FUNCTION_BLOCK TestingSequence1 (* Composite Function Block Type *)
  (* Standard: 61499-2 *)
  (* Version 0.0, 7/2/2026, template *)
  PACKAGE Main;
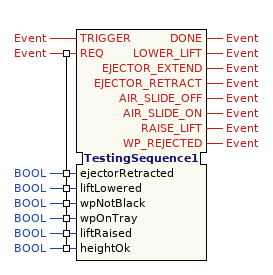
  EVENT_INPUT
    TRIGGER; (* Initialization Request *)
    REQ WITH ejectorRetracted, liftLowered, wpNotBlack, wpOnTray, liftRaised, heightOk; (* Normal Execution Request *)
  END_EVENT
  EVENT_OUTPUT
    DONE; (* Initialization Confirm *)
    LOWER_LIFT; (* Execution Confirmation *)
    EJECTOR_EXTEND;
    EJECTOR_RETRACT;
    AIR_SLIDE_OFF;
    AIR_SLIDE_ON;
    RAISE_LIFT;
    WP_REJECTED;
  END_EVENT
  VAR_INPUT
    ejectorRetracted : BOOL; (* Input event qualifier *)
    liftLowered : BOOL;
    wpNotBlack : BOOL;
    wpOnTray : BOOL;
    liftRaised : BOOL;
    heightOk : BOOL;
  END_VAR
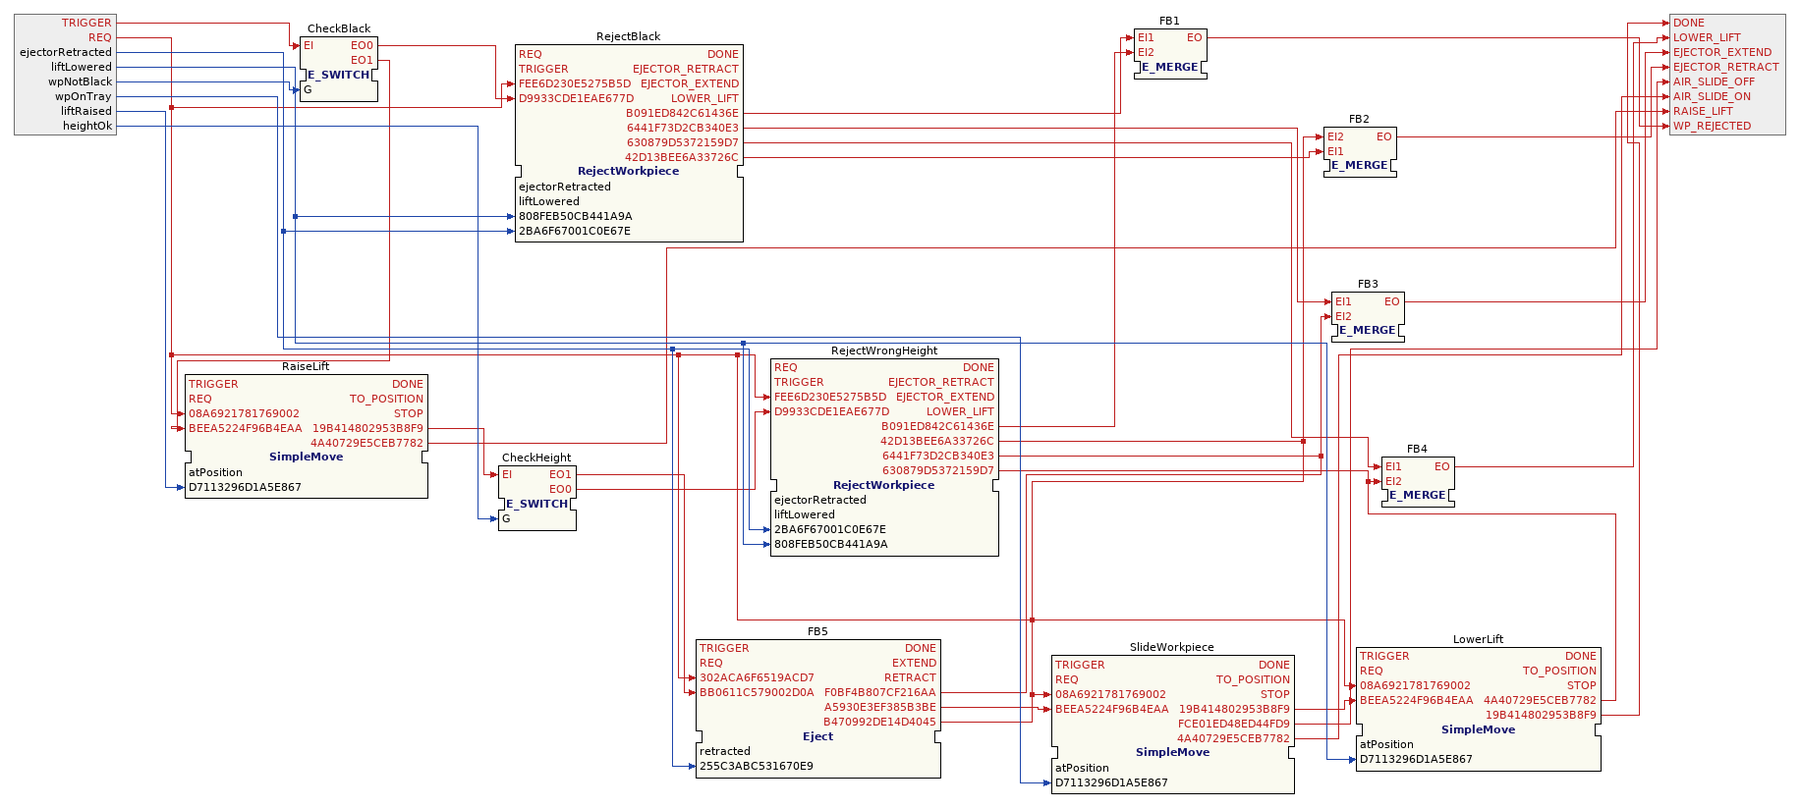
  FBS
    CheckBlack : E_SWITCH;
    RejectBlack : RejectWorkpiece;
    RaiseLift : SimpleMove;
    CheckHeight : E_SWITCH;
    RejectWrongHeight : RejectWorkpiece;
    FB1 : E_MERGE;
    FB2 : E_MERGE;
    FB3 : E_MERGE;
    FB4 : E_MERGE;
    FB5 : Eject;
    SlideWorkpiece : SimpleMove;
    LowerLift : SimpleMove;
  END_FBS
  EVENT_CONNECTIONS
    TRIGGER TO CheckBlack.EI;
    REQ TO RejectBlack.FEE6D230E5275B5D;
    REQ TO RaiseLift.08A6921781769002;
    REQ TO FB5.302ACA6F6519ACD7;
    REQ TO RejectWrongHeight.FEE6D230E5275B5D;
    REQ TO SlideWorkpiece.08A6921781769002;
    REQ TO LowerLift.08A6921781769002;
    CheckBlack.EO0 TO RejectBlack.D9933CDE1EAE677D;
    CheckBlack.EO1 TO RaiseLift.BEEA5224F96B4EAA;
    RaiseLift.19B414802953B8F9 TO CheckHeight.EI;
    CheckHeight.EO1 TO FB5.BB0611C579002D0A;
    CheckHeight.EO0 TO RejectWrongHeight.D9933CDE1EAE677D;
    RaiseLift.4A40729E5CEB7782 TO RAISE_LIFT;
    RejectBlack.B091ED842C61436E TO FB1.EI1;
    RejectBlack.6441F73D2CB340E3 TO FB3.EI1;
    RejectBlack.630879D5372159D7 TO FB4.EI1;
    RejectWrongHeight.B091ED842C61436E TO FB1.EI2;
    RejectWrongHeight.42D13BEE6A33726C TO FB2.EI2;
    RejectBlack.42D13BEE6A33726C TO FB2.EI1;
    FB2.EO TO EJECTOR_RETRACT;
    FB1.EO TO WP_REJECTED;
    FB3.EO TO EJECTOR_EXTEND;
    FB5.F0BF4B807CF216AA TO FB3.EI2;
    RejectWrongHeight.6441F73D2CB340E3 TO FB3.EI2;
    RejectWrongHeight.630879D5372159D7 TO FB4.EI2;
    FB4.EO TO LOWER_LIFT;
    SlideWorkpiece.19B414802953B8F9 TO LowerLift.BEEA5224F96B4EAA;
    FB5.A5930E3EF385B3BE TO SlideWorkpiece.BEEA5224F96B4EAA;
    FB5.B470992DE14D4045 TO FB2.EI2;
    FB5.B470992DE14D4045 TO SlideWorkpiece.08A6921781769002;
    SlideWorkpiece.FCE01ED48ED44FD9 TO AIR_SLIDE_OFF;
    SlideWorkpiece.4A40729E5CEB7782 TO AIR_SLIDE_ON;
    LowerLift.4A40729E5CEB7782 TO FB4.EI2;
    LowerLift.19B414802953B8F9 TO DONE;
  END_CONNECTIONS
  DATA_CONNECTIONS
    heightOk TO CheckHeight.G;
    liftRaised TO RaiseLift.D7113296D1A5E867;
    liftLowered TO RejectBlack.808FEB50CB441A9A;
    ejectorRetracted TO RejectBlack.2BA6F67001C0E67E;
    wpNotBlack TO CheckBlack.G;
    ejectorRetracted TO FB5.255C3ABC531670E9;
    ejectorRetracted TO RejectWrongHeight.2BA6F67001C0E67E;
    liftLowered TO LowerLift.D7113296D1A5E867;
    liftLowered TO RejectWrongHeight.808FEB50CB441A9A;
    wpOnTray TO SlideWorkpiece.D7113296D1A5E867;
  END_CONNECTIONS
END_FUNCTION_BLOCK
